(* CoDeSys 2.3 export: ld.exp *)

(* POU PLC_LD_PRG_TR, LD *)
PROGRAM PLC_LD_PRG_TR
VAR
END_VAR
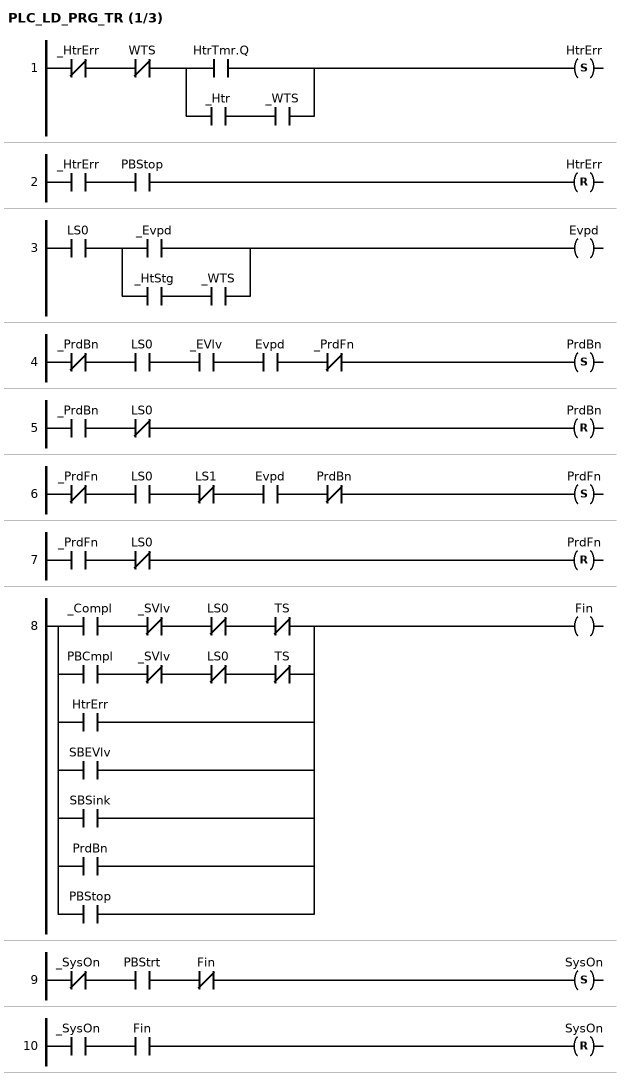
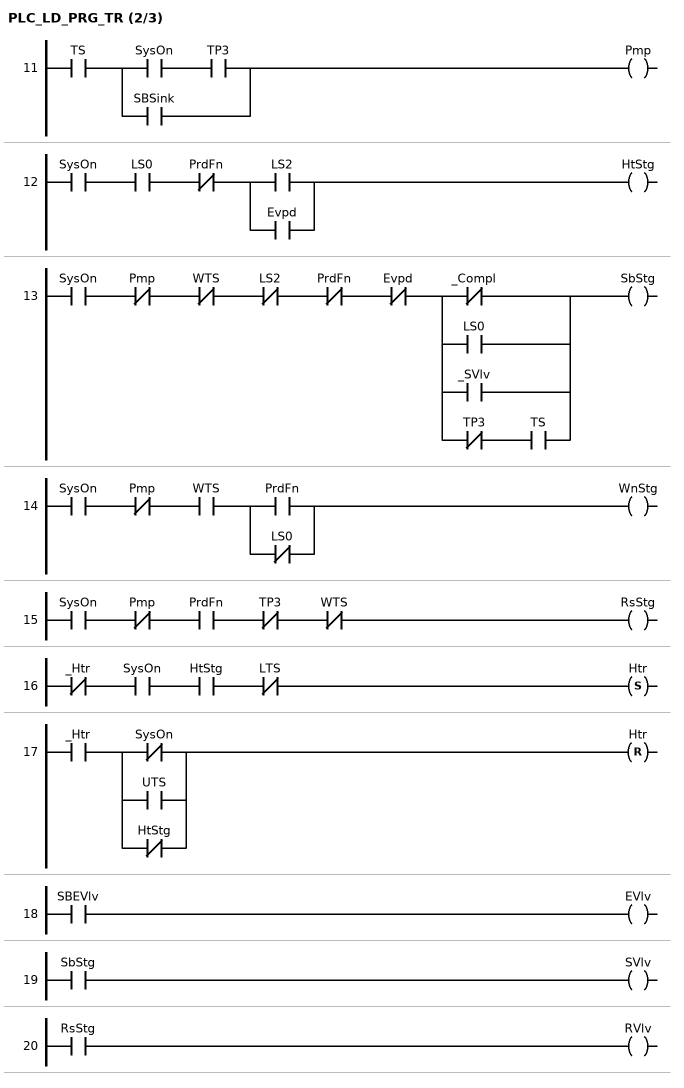
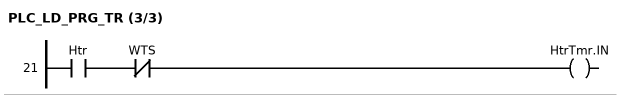
_LD_ (* Ladder Diagram *)
NETWORK 1
	[/_HtrErr] - [/WTS] - { [HtrTmr.Q] | [_Htr] - [_WTS] } --- (S HtrErr)
NETWORK 2
	[_HtrErr] - [PBStop] --- (R HtrErr)
NETWORK 3
	[LS0] - { [_Evpd] | [_HtStg] - [_WTS] } --- (Evpd)
NETWORK 4
	[/_PrdBn] - [LS0] - [_EVlv] - [Evpd] - [/_PrdFn] --- (S PrdBn)
NETWORK 5
	[_PrdBn] - [/LS0] --- (R PrdBn)
NETWORK 6
	[/_PrdFn] - [LS0] - [/LS1] - [Evpd] - [/PrdBn] --- (S PrdFn)
NETWORK 7
	[_PrdFn] - [/LS0] --- (R PrdFn)
NETWORK 8
	{ [_Compl] - [/_SVlv] - [/LS0] - [/TS] | [PBCmpl] - [/_SVlv] - [/LS0] - [/TS] | [HtrErr] | [SBEVlv] | [SBSink] | [PrdBn] | [PBStop] } --- (Fin)
NETWORK 9
	[/_SysOn] - [PBStrt] - [/Fin] --- (S SysOn)
NETWORK 10
	[_SysOn] - [Fin] --- (R SysOn)
NETWORK 11
	[TS] - { [SysOn] - [TP3] | [SBSink] } --- (Pmp)
NETWORK 12
	[SysOn] - [LS0] - [/PrdFn] - { [LS2] | [Evpd] } --- (HtStg)
NETWORK 13
	[SysOn] - [/Pmp] - [/WTS] - [/LS2] - [/PrdFn] - [/Evpd] - { [/_Compl] | [LS0] | [_SVlv] | [/TP3] - [TS] } --- (SbStg)
NETWORK 14
	[SysOn] - [/Pmp] - [WTS] - { [PrdFn] | [/LS0] } --- (WnStg)
NETWORK 15
	[SysOn] - [/Pmp] - [PrdFn] - [/TP3] - [/WTS] --- (RsStg)
NETWORK 16
	[/_Htr] - [SysOn] - [HtStg] - [/LTS] --- (S Htr)
NETWORK 17
	[_Htr] - { [/SysOn] | [UTS] | [/HtStg] } --- (R Htr)
NETWORK 18
	[SBEVlv] --- (EVlv)
NETWORK 19
	[SbStg] --- (SVlv)
NETWORK 20
	[RsStg] --- (RVlv)
NETWORK 21
	[Htr] - [/WTS] --- (HtrTmr.IN)
_END_LD_
(* the same logic as Structured Text *)
(* Network 1 *)
IF NOT _HtrErr AND NOT WTS AND (HtrTmr.Q OR _Htr AND _WTS) THEN HtrErr := TRUE; END_IF;
(* Network 2 *)
IF _HtrErr AND PBStop THEN HtrErr := FALSE; END_IF;
(* Network 3 *)
Evpd := LS0 AND (_Evpd OR _HtStg AND _WTS);
(* Network 4 *)
IF NOT _PrdBn AND LS0 AND _EVlv AND Evpd AND NOT _PrdFn THEN PrdBn := TRUE; END_IF;
(* Network 5 *)
IF _PrdBn AND NOT LS0 THEN PrdBn := FALSE; END_IF;
(* Network 6 *)
IF NOT _PrdFn AND LS0 AND NOT LS1 AND Evpd AND NOT PrdBn THEN PrdFn := TRUE; END_IF;
(* Network 7 *)
IF _PrdFn AND NOT LS0 THEN PrdFn := FALSE; END_IF;
(* Network 8 *)
Fin := _Compl AND NOT _SVlv AND NOT LS0 AND NOT TS OR PBCmpl AND NOT _SVlv AND NOT LS0 AND NOT TS OR HtrErr OR SBEVlv OR SBSink OR PrdBn OR PBStop;
(* Network 9 *)
IF NOT _SysOn AND PBStrt AND NOT Fin THEN SysOn := TRUE; END_IF;
(* Network 10 *)
IF _SysOn AND Fin THEN SysOn := FALSE; END_IF;
(* Network 11 *)
Pmp := TS AND (SysOn AND TP3 OR SBSink);
(* Network 12 *)
HtStg := SysOn AND LS0 AND NOT PrdFn AND (LS2 OR Evpd);
(* Network 13 *)
SbStg := SysOn AND NOT Pmp AND NOT WTS AND NOT LS2 AND NOT PrdFn AND NOT Evpd AND (NOT _Compl OR LS0 OR _SVlv OR NOT TP3 AND TS);
(* Network 14 *)
WnStg := SysOn AND NOT Pmp AND WTS AND (PrdFn OR NOT LS0);
(* Network 15 *)
RsStg := SysOn AND NOT Pmp AND PrdFn AND NOT TP3 AND NOT WTS;
(* Network 16 *)
IF NOT _Htr AND SysOn AND HtStg AND NOT LTS THEN Htr := TRUE; END_IF;
(* Network 17 *)
IF _Htr AND (NOT SysOn OR UTS OR NOT HtStg) THEN Htr := FALSE; END_IF;
(* Network 18 *)
EVlv := SBEVlv;
(* Network 19 *)
SVlv := SbStg;
(* Network 20 *)
RVlv := RsStg;
(* Network 21 *)
HtrTmr.IN := Htr AND NOT WTS;
END_PROGRAM
